(* IEC 61131-3 sources: rtacc/examples/ST, 1 file *)

(* ---- invert.st ---- *)
FUNCTION NotBool : BOOL
VAR_INPUT
    x : BOOL;
END_VAR

NotBool := NOT x;

END_FUNCTION
